Staubli VAL3: setjointmode.pgx

public program setjointmode()
  local num l_i
begin
  $jogMode(1)
   for l_i = 0 to size(sShowType)-1
    sShowType[l_i]=sJoint[l_i]
  endFor
end
